(* IEC 61131-3 sources: codesys-framework/txt/application/ToDo/Utils/Moving Average/Impl/FB_ExponentialMovingAverage, 3 files *)

(* ---- AddValue.method.st ---- *)
METHOD AddValue
VAR_INPUT
	lrValue 	: LREAL;
END_VAR
VAR
	lrMultiplier 	: LREAL;
END_VAR

// --- BEGIN IMPLEMENTATION ---

lrMultiplier := 2.0 / UINT_TO_LREAL(_scSysPar.iNbrOfItemsForAverage + 1);

IF _lrEma = 0 THEN
	_lrEma := lrValue;
	RETURN;
END_IF

_lrEma := (lrValue * lrMultiplier) + (_lrEma * (1 - lrMultiplier));

(* ---- Reset.method.st ---- *)
METHOD Reset
VAR_INPUT
END_VAR
VAR
	i 	: UINT;
END_VAR

// --- BEGIN IMPLEMENTATION ---

_lrEma := 0;

(* ---- SysPar.prop.st ---- *)
PROPERTY SysPar : SC_SystemParametersMovingAverage

// --- BEGIN IMPLEMENTATION ---

// ----------- SET -----------
VAR
END_VAR

// -- BEGIN IMPLEMENTATION SET --
_scSysPar := SysPar;
